(* IEC 61131-3 sources: volt/packages/volt-lsp-iec/test-corpus/bakon-nano/Device/Plc Logic/Application/Library Manager/NetVarUdp, 22 files *)

(* ---- CLIENT_ACCEPT.dut ---- *)
TYPE CLIENT_ACCEPT :
STRUCT
	DISOCKET : DINT;
	STIPADDRESS : STRING(20);
END_STRUCT
END_TYPE

(* ---- CLIENT_REPLY.dut ---- *)
TYPE CLIENT_REPLY :
STRUCT
	DIBYTESRECEIVED : __XINT;
	DWIPADDRESS : DWORD;
	STIPADDRESSTRANSMITTER : STRING;
END_STRUCT
END_TYPE

(* ---- NETVARDATAITEM_UDP.dut ---- *)
TYPE NETVARDATAITEM_UDP :
STRUCT
	PADDRESS : POINTER TO BYTE;
	NDATALEN : INT;
	SITYPE : SINT := -1;
END_STRUCT
END_TYPE

(* ---- NETVAROD_SERVICE_UDP.dut ---- *)
TYPE NETVAROD_SERVICE_UDP :
(
	ODSTATEFREE := 0,
	ODREADREQUEST,
	ODREADREQUESTREPLY,
	ODWRITEREQUEST,
	ODWRITEREQUESTREPLY,
	ODACKNOWLEDGEMENT,
	ODBOOTUPREQUEST,
	ODERRORREPLYUNNOWN := 20,
	ODERRORREPLYITEMS,
	ODERRORREPLYACCESS,
	ODERRORREPLYIDX,
	ODERRORREPLYSUB,
	ODERRORREPLYLEN,
	ODERRORWRONGSERVICE,
	ODERRORTIMEOUT,
	ODERRORREPLYCPUSTOPPED,
	ODERRORDATALENGTH,
	ODSTATEBUSY := 100
);
END_TYPE

(* ---- NETVARTELEGRAMM_UDP.dut ---- *)
TYPE NETVARTELEGRAMM_UDP :
STRUCT
	HEADER : NetVarTlgHeader_Udp;
	PDATA : ARRAY [0..(Parameters.UdpPacketSize - 1)] OF BYTE;
END_STRUCT
END_TYPE

(* ---- NETVARTLGHEADER_UDP.dut ---- *)
TYPE NETVARTLGHEADER_UDP :
STRUCT
	DWIDENTITY : DWORD := 16#33532D00;
	DWID : DWORD;
	NINDEX : INT;
	NSUBINDEX : INT;
	NITEMS : INT;
	NLEN : INT;
	NCOUNTER : INT;
	BYFLAGS : BYTE;
	BYCHECKSUM : BYTE;
END_STRUCT
END_TYPE

(* ---- NETVARUDPDIAGSTRUCT.dut ---- *)
TYPE NETVARUDPDIAGSTRUCT :
STRUCT
	NSENDCOUNT : UDINT;
	TLASTSEND : TIME;
	NRECEIVECOUNT : UDINT;
	TLASTRECEIVE : TIME;
	NWRITECOUNT : UDINT;
	SLASTERROR : NetVarUDPError;
	TLASTERROR : TIME;
	NERRORCOUNT : UINT;
	NACKNOWLEDGES : UINT;
	BSENDERSTOPPED : BOOL;
END_STRUCT
END_TYPE

(* ---- NETVARUDPERROR.dut ---- *)
TYPE NETVARUDPERROR :
(
	NETVARUDPERROR_NOERROR := 0,
	NETVARUDPERROR_UDPSENDDATA,
	NETVARUDPERROR_UDPSENDACKN,
	NETVARUDPERROR_NOACKNOWLEDGEMENT,
	NETVARUDPERROR_NOTACKNOWLEDGED,
	NETVARUDPERROR_UDPSENDBOOTUPREQUEST,
	NETVARUDPERROR_UDPANSWERBOOTUPREQUEST,
	NETVARUDPERROR_CHECKSUM,
	NETVARUDPERROR_LAYOUT,
	NETVARUDPERROR_PACKETSIZEMISMATCH,
	NETVARUDPERROR_UDPNETWORKMANAGER_NOT_READY := 20,
	NETVARUDPERROR_UNKNOWN := 100
);
END_TYPE

(* ---- GLOBALE_VARIABLEN.gvl ---- *)
VAR_GLOBAL
	G_BCPUSTOPNETVAR : BOOL;
	TELEGRAM_IDENT : DWORD := 16#33532D00;
END_VAR

(* ---- PARAMETERS.gvl ---- *)
VAR_GLOBAL
	UDPPACKETSIZE : UINT := 256;
END_VAR

(* ---- CALLBACKNETVAR.pou ---- *)
FUNCTION CALLBACKNETVAR : BYTE
VAR_INPUT
	DWEVENT : DWORD;
	DWFILTER : DWORD;
	DWOWNER : DWORD;
END_VAR
END_FUNCTION

(* ---- CALLBACKTASKCODENC.pou ---- *)
FUNCTION CALLBACKTASKCODENC : BYTE
VAR_INPUT
	DWEVENT : DWORD;
	DWFILTER : DWORD;
	DWOWNER : DWORD;
END_VAR
END_FUNCTION

(* ---- GETIPADDRESS.pou ---- *)
FUNCTION GETIPADDRESS : UDINT
VAR_INPUT
	STIPADDRESS : STRING;
END_VAR
END_FUNCTION

(* ---- SWAP.pou ---- *)
FUNCTION SWAP : BOOL
VAR_INPUT
	BSWAP : BOOL;
	PI : POINTER TO BYTE;
	NSIZE : INT;
END_VAR
END_FUNCTION

(* ---- UDPGETRECEIVEDATASIZE.pou ---- *)
FUNCTION UDPGETRECEIVEDATASIZE : DINT
VAR_INPUT
	HSOCKET : RTS_IEC_HANDLE;
END_VAR
END_FUNCTION

(* ---- UDPOPENRECEIVESOCKET.pou ---- *)
FUNCTION UDPOPENRECEIVESOCKET : RTS_IEC_HANDLE
VAR_INPUT
	IPORT : INT;
END_VAR
END_FUNCTION

(* ---- UDPOPENSENDSOCKET.pou ---- *)
FUNCTION UDPOPENSENDSOCKET : RTS_IEC_HANDLE
VAR_INPUT
	IPORT : INT;
END_VAR
END_FUNCTION

(* ---- UDPRECEIVEDATA.pou ---- *)
FUNCTION UDPRECEIVEDATA : CLIENT_REPLY
VAR_INPUT
	HSOCKET : RTS_IEC_HANDLE;
	IPORT : INT;
	PBYDATA : POINTER TO BYTE;
	DIDATASIZE : __XINT;
END_VAR
END_FUNCTION

(* ---- UDPSENDDATA.pou ---- *)
FUNCTION UDPSENDDATA : __XINT
VAR_INPUT
	HSOCKET : RTS_IEC_HANDLE;
	IPORT : INT;
	STIPADDRESS : STRING;
	PBYDATA : POINTER TO BYTE;
	DIDATASIZE : DINT;
END_VAR
END_FUNCTION

(* ---- NETVARMANAGER_UDP_FB.pou ---- *)
FUNCTION_BLOCK NETVARMANAGER_UDP_FB
VAR_INPUT
	NNETVARPDO_RX : INT;
	PNETVARPDO_RX : POINTER TO NetVarPDO_Rx_Udp;
	NNETVARPDO_TX : INT;
	PNETVARPDO_TX : POINTER TO NetVarPDO_Tx_Udp;
	BBYTESWAP : BOOL;
	DWIDENTITY : DWORD;
	INEWTLGPERCYCLE : INT := 0;
	UIPACKETSIZE : UINT := Parameters.UdpPacketSize;
	IPORT : INT := 1202;
END_VAR
VAR
	HSOKETRX : RTS_IEC_HANDLE := RTS_INVALID_HANDLE;
	HSOKETTX : RTS_IEC_HANDLE := RTS_INVALID_HANDLE;
	DIRXLEN : DINT;
	DIOFFSET : __XINT;
	DICALLCOUNTER : DINT;
	DIMSGCOUNTER : DINT := 0;
	DWONEIPADDRESS : DWORD;
	PSZHOSTNAME : STRING(80);
	READ : CLIENT_REPLY;
	TLG : NetVarTelegramm_Udp;
	TLGTEMP : NetVarTelegramm_Udp;
	NSTATUS : INT;
	N : INT;
	BISACTIV : BOOL;
	BREADNEXT : BOOL;
	BTLGREADY : BOOL;
	ITLGPERCYCLE : INT;
	ITLGCOUNT : INT;
	TINHIBIT : TON := STRUCT(pt := TIME#1s500ms);
	RESULT : RTS_IEC_RESULT;
	HOST : SOCK_HOSTENT;
	ILEN : INT;
	BACKNOWLEDGENEEDED : BOOL := FALSE;
	BRECEIVESOCKETOPENED : BOOL := TRUE;
	PAPPCURRENT : POINTER TO APPLICATION;
	DWRESULT : DWORD;
	HEVENTSTOP : __XWORD;
	HINTERFACESTOP : __XWORD;
	ITF : ICmpEventCallback;
	BPREPARESTOP : BOOL;
	HEVENTSTOPDONE : __XWORD;
	HINTERFACESTOPDONE : __XWORD;
	HEVENTDEBUGLOOP : __XWORD;
	HINTERFACEDEBUGLOOP : __XWORD;
END_VAR
END_FUNCTION_BLOCK

METHOD CLOSESOCKETS
END_METHOD

METHOD EVENTCALLBACK : UDINT
VAR_INPUT
	PEVENTPARAM : POINTER TO EventParam;
END_VAR
END_METHOD

METHOD FB_EXIT : BOOL
VAR_INPUT
	BINCOPYCODE : BOOL;
END_VAR
END_METHOD

METHOD NETVARGETCONNECTSTATUS_UDP : BOOL
VAR_INPUT
	NBASISID : INT;
END_VAR
VAR_OUTPUT
	BCONNECTNEWDATA : BOOL;
	BCONNECTERROR : BOOL;
	DWERRORCODE : DWORD;
END_VAR
END_METHOD

METHOD REGISTEREVENTS : BOOL
END_METHOD

METHOD SEND : BOOL
END_METHOD

METHOD SETPACKETSIZEMISMATCHERROR : BOOL
END_METHOD

METHOD UNREGISTEREVENTS
END_METHOD

(* ---- NETVARPDO_RX_UDP.pou ---- *)
FUNCTION_BLOCK NETVARPDO_RX_UDP
VAR_INPUT
	SNETTELEGRAMM : NetVarTelegramm_UDP;
	TIMEOUT : TON := STRUCT(PT := TIME#500ms);
	BNEWMESSAGE : BOOL;
	NINDEX : INT := -1;
	NSUBINDEX : INT := -1;
	DIBYTESSEND : DINT;
	BRECEIVED : BOOL := FALSE;
	BACTIVE : BOOL := TRUE;
	PDATAITEMS : POINTER TO NetVarDataItem_UDP;
	WDRVNR : WORD;
	NDATAITEMS : INT := -1;
	BYCHECKSUM : BYTE;
	BREQUESTATBOOTUP : BOOL := TRUE;
	STIPADDRESSTRANSMITTER : STRING(20);
	PNETVARMANAGER_UDP : POINTER TO NetVarManager_Udp_FB;
	PNETVARPDO_RX_DIAGNOSIS : POINTER TO NetVarUDPDiagStruct;
	STIPADDRESSBROADCAST : STRING(20);
END_VAR
VAR_OUTPUT
	NSTATUS : INT;
	BDATANEW : BOOL;
END_VAR
VAR
	PPTRTOPDO_TXDATA : POINTER TO ARRAY [0..127] OF BYTE;
	PPTRTODATA : POINTER TO ARRAY [0..127] OF BYTE;
	DATAITEM : NetVarDataItem_UDP;
	I : INT;
	N : INT;
	NLEN : INT;
	NDESTIX : INT;
	NDESTORDER : INT;
	IDATAIX : INT;
	NLASTRXCOUNTER : INT;
	BINIT : BOOL := TRUE;
	BCHECKSUMVALID : BOOL := TRUE;
	SITYPE : SINT := -1;
END_VAR
END_FUNCTION_BLOCK

METHOD NEWDATAREC
END_METHOD

METHOD SETERROR : BOOL
VAR_INPUT
	ERROR : NetVarUDPError;
END_VAR
END_METHOD

(* ---- NETVARPDO_TX_UDP.pou ---- *)
FUNCTION_BLOCK NETVARPDO_TX_UDP
VAR_INPUT
	NDATAITEMS : INT := -1;
	PDATAITEMS : POINTER TO NetVarDataItem_Udp;
	WDRVNR : WORD;
	NINDEX : INT := -1;
	NSUBINDEX : INT := -1;
	BWITHCHECKSUM : BOOL;
	BYCHECKSUM : BYTE;
	BWITHACKNOWLEDGE : BOOL;
	PBEXPRESSION : POINTER TO BOOL;
	BANSWERBOOTUPREQUEST : BOOL := TRUE;
	BBOOTUPREQUESTRECEIVED : BOOL;
	INHIBITTIMER : TON := STRUCT(PT := TIME#100ms);
	REPEATTIMER : TON := STRUCT(PT := TIME#500ms);
	STIPADDRESSBOOTUPREQUEST : STRING(20);
	SNETTELEGRAMM : NetVarTelegramm_UDP;
	BACTIVE : BOOL := TRUE;
	PNETVARMANAGER_UDP : POINTER TO NetVarManager_Udp_FB;
	PNETVARPDO_TX_DIAGNOSIS : POINTER TO NetVarUDPDiagStruct;
	BBEFOREAPPLICATION : BOOL := FALSE;
	STIPADDRESSBROADCAST : STRING(20);
END_VAR
VAR_OUTPUT
	NSTATUS : INT;
END_VAR
VAR
	DIBYTESSEND : __XINT;
	DATAITEM : NetVarDataItem_UDP;
	I : INT;
	N : INT;
	NLEN : INT;
	NDESTIX : INT;
	NDESTORDER : INT;
	IDATAIX : INT;
	NLENTOSEND : INT;
	BSEND : BOOL := TRUE;
	BSENDHARD : BOOL;
	BINIT : BOOL := TRUE;
	BACKNEXPECTED : BOOL := FALSE;
	STLGBOOTUPREQ : NetVarTelegramm_UDP;
	BEXPR : BOOL := FALSE;
	SITYPE : SINT := -1;
END_VAR
END_FUNCTION_BLOCK

METHOD ACKNOWLEDGE : BOOL
END_METHOD

METHOD PDO_TXSENDHARD
END_METHOD

METHOD SETERROR : BOOL
VAR_INPUT
	ERROR : NetVarUDPError;
END_VAR
END_METHOD
